(* PLC project g_guard_lock_no_rundown, Anonymous Benchmark Suite 1.0 *)
(* stored: creationDateTime 2026-08-28T00:00:00 *)

PROGRAM g_guard_lock_no_rundown
  VAR_INPUT
    OpenReq : BOOL;
    DoorClosed : BOOL;
    RunCmd : BOOL;
  END_VAR
  VAR_OUTPUT
    Motor : BOOL;
    Unlocked : BOOL;
  END_VAR

(* LD diagram, written out as Structured Text *)
Unlocked := OpenReq;
Motor := RunCmd AND DoorClosed AND NOT OpenReq;
END_PROGRAM

CONFIGURATION Config0
  RESOURCE Res0 ON PLC
    TASK tcyclic(INTERVAL := T#10ms, PRIORITY := 0);
    PROGRAM inst0 WITH tcyclic : g_guard_lock_no_rundown;
  END_RESOURCE
END_CONFIGURATION
